// TIA Portal V20 export
FUNCTION_BLOCK "OVLADANI_LASER"   // FB400, LAD
{ S7_Optimized_Access := 'TRUE' }
// stored: AutoNumber false, MemoryReserve 100, SetENOAutomatically false
   VAR
      SQCR : Int;
      SQCR_WHILE : Int;
      SET_WHILE : Bool;
      NAZEV_PROGRAMU : String[20];
      DELKA_STRINGU : Int;
      CHAR_K_ZAPISU : Array[0..71] of Char;
   END_VAR
   VAR CONSTANT
      STEP_0 : Int := 0;
      STEP_5 : Int := 5;
      STEP_10 : Int := 10;
      STEP_15 : Int := 15;
      STEP_20 : Int := 20;
      STEP_25 : Int := 25;
      STEP_30 : Int := 30;
      STEP_35 : Int := 35;
      STEP_40 : Int := 40;
      STEP_45 : Int := 45;
      STEP_50 : Int := 50;
      STEP_55 : Int := 55;
      STEP_60 : Int := 60;
      STEP_65 : Int := 65;
      STEP_70 : Int := 70;
      STEP_75 : Int := 75;
      STEP_80 : Int := 80;
      STEP_85 : Int := 85;
      STEP_90 : Int := 90;
      STEP_95 : Int := 95;
      STEP_100 : Int := 100;
   END_VAR
BEGIN

REGION Network 1
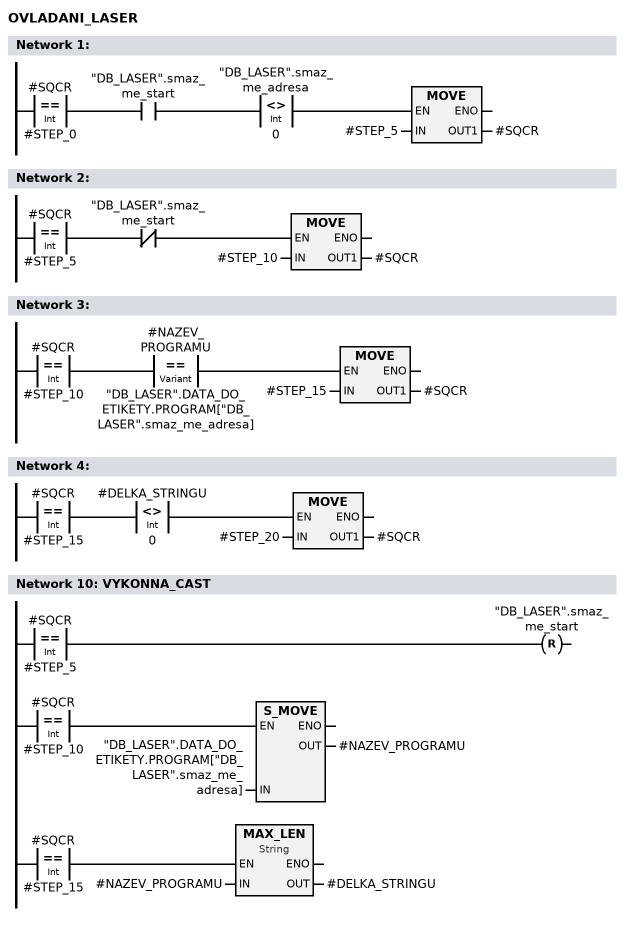
   RUNG wire#powerrail
      { S7_Templates := "SrcType := Int" } EQ_Contact(in1 := #SQCR, in2 := #STEP_0)
      Contact( "DB_LASER".smaz_me_start )
      { S7_Templates := "SrcType := Int" } NE_Contact(in1 := "DB_LASER".smaz_me_adresa, in2 := 0)
      Move(in := #STEP_5, out1 => #SQCR)
   END_RUNG
   // the same network as SCL:
   IF (#SQCR = #STEP_0) AND "DB_LASER".smaz_me_start AND ("DB_LASER".smaz_me_adresa <> 0) THEN
       #SQCR := #STEP_5;
   END_IF;
END_REGION

REGION Network 2
   RUNG wire#powerrail
      { S7_Templates := "SrcType := Int" } EQ_Contact(in1 := #SQCR, in2 := #STEP_5)
      I_Contact( "DB_LASER".smaz_me_start )
      Move(in := #STEP_10, out1 => #SQCR)
   END_RUNG
   // the same network as SCL:
   IF (#SQCR = #STEP_5) AND NOT "DB_LASER".smaz_me_start THEN #SQCR := #STEP_10; END_IF;
END_REGION

REGION Network 3
   RUNG wire#powerrail
      { S7_Templates := "SrcType := Int" } EQ_Contact(in1 := #SQCR, in2 := #STEP_10)
      { S7_Templates := "SrcType := Variant" } EQ_Contact(in1 := #NAZEV_PROGRAMU, in2 := "DB_LASER".DATA_DO_ETIKETY.PROGRAM["DB_LASER".smaz_me_adresa])
      Move(in := #STEP_15, out1 => #SQCR)
   END_RUNG
   // the same network as SCL:
   IF (#SQCR = #STEP_10) AND (#NAZEV_PROGRAMU = "DB_LASER".DATA_DO_ETIKETY.PROGRAM["DB_LASER".smaz_me_adresa]) THEN
       #SQCR := #STEP_15;
   END_IF;
END_REGION

REGION Network 4
   RUNG wire#powerrail
      { S7_Templates := "SrcType := Int" } EQ_Contact(in1 := #SQCR, in2 := #STEP_15)
      { S7_Templates := "SrcType := Int" } NE_Contact(in1 := #DELKA_STRINGU, in2 := 0)
      Move(in := #STEP_20, out1 => #SQCR)
   END_RUNG
   // the same network as SCL:
   IF (#SQCR = #STEP_15) AND (#DELKA_STRINGU <> 0) THEN #SQCR := #STEP_20; END_IF;
END_REGION

REGION Network 5: STEP_20 SCL NETVORK X
END_REGION

REGION Network 10: VYKONNA_CAST
   IF #SQCR = #STEP_5 THEN "DB_LASER".smaz_me_start := FALSE; END_IF;
   IF #SQCR = #STEP_10 THEN
       #NAZEV_PROGRAMU := "DB_LASER".DATA_DO_ETIKETY.PROGRAM["DB_LASER".smaz_me_adresa];
   END_IF;
   IF #SQCR = #STEP_15 THEN MAX_LEN(in := #NAZEV_PROGRAMU, out => #DELKA_STRINGU); END_IF;
END_REGION

REGION Network 12 (SCL)
   IF #SQCR = #STEP_20 THEN
       // zapsani počátečního znaku 
       #CHAR_K_ZAPISU[0] := "DB_LASER".DATA_DO_DAT.ZAVORKA_P;



       // vytvoření prdelky k názvu programu z laseru
       #CHAR_K_ZAPISU[#DELKA_STRINGU + 1] := "DB_LASER".DATA_DO_DAT.XLP[0];
       #CHAR_K_ZAPISU[#DELKA_STRINGU + 2] := "DB_LASER".DATA_DO_DAT.XLP[1];
       #CHAR_K_ZAPISU[#DELKA_STRINGU + 3] := "DB_LASER".DATA_DO_DAT.XLP[2];
       #CHAR_K_ZAPISU[#DELKA_STRINGU + 4] := "DB_LASER".DATA_DO_DAT.XLP[3];
       #CHAR_K_ZAPISU[#DELKA_STRINGU + 5] := "DB_LASER".DATA_DO_DAT.ZAVORKA_P;

       // dinamický zápis názvu podle délky stringu 
       WHILE #SET_WHILE DO
           IF #SQCR_WHILE > #DELKA_STRINGU THEN
               #SQCR_WHILE := 0;
               #SET_WHILE := FALSE;
               #SQCR := #STEP_25;
           ELSE
               #SQCR_WHILE := #SQCR_WHILE + 1;
           END_IF;
           #CHAR_K_ZAPISU[#SQCR_WHILE + 1] := #NAZEV_PROGRAMU[#SQCR_WHILE];
       END_WHILE;

   END_IF;
END_REGION
END_FUNCTION_BLOCK
